INTERFACE I_Clock EXTENDS __SYSTEM.IQueryInterface

PROPERTY Now : LTIME
GET
END_GET
END_PROPERTY

END_INTERFACE

(* stored: Version 1.1.0.1
   Itf I_Clock: Id {82fe060f-c53c-4bbf-9d7d-8a13a7ae689c}
   Property Now: Id {64bc7d1c-0305-48dd-b2f7-c6380cba35e1}
   Get Get: Id {e52e276b-2515-40ca-bd51-3730fee8b880} *)
